Universal Robots PolyScope program: P1140 INVITE_Demo_1111.urp

Program P1140 INVITE_Demo_1111 (installation=default_INVITE directory=/programs createdIn=5.10.1 lastSavedIn=5.23.0 robotSerialNumber=20245590068)
Calibrated DH parameters: a=[0.00013, -0.03651, -0.389144, 0.000102, 0.000008, 0]; d=[0.162613, 192.230671, -179.915756, -12.181517, 0.099698, 0.099535]; alpha=[1.57038, 0.002205, 0.004138, 1.570804, -1.571025, 0]; deltaTheta=[-0.000001, 1.484886, 4.928506, -0.130209, 0, 0]
InitVariablesNode variables(variable(name=AMR_Position, expression=struct(position_identifier=0, x1=0, x2=0, y1=0, y2=0, theta1=0, theta2=0)), variable(name=CAM_Pose, expression=p[0,0,0,0,0,0]), variable(name=CAM_Relation, expression=""), variable(name=CMD_Abort, expression=False), variable(name=CMD_Clear, expression=False), variable(name=CMD_Reset, expression=False), variable(name=CMD_Start, expression=False), variable(name=CMD_Suspend, expression=False), variable(name=CMD_Unhold, expression=False), variable(name=CMD_Unsuspend, expression=False), variable(name=CNT_Rack_Output, expression=0), variable(name=FNC_Freedrive, expression=False), variable(name=PRC_TubCounter, expression=0), variable(name=PRC_TubNumber, expression=0), variable(name=STP, expression=0), variable(name=TMR_Barcode, expression=0), variable(name=easyPickCount, expression=0), variable(name=easyPickCount_5, expression=0), variable(name=easyPickNoObj, expression=0), variable(name=easyPickNoObj_5, expression=0), variable(name=easyPickParts, expression=0), variable(name=easyPickParts_5, expression=0))
BeforeStart
  Folder Scripts [hidden by the author, left out]
  Folder BeforeStarts [hidden by the author, left out]
  Script file /programs/04 Scripts/krish.script
    | def vibration_2():
    | 	set_analog_out(0,0.4)
    | 	sleep(0.8)
    | 	set_analog_out(0,0.0)
    | 	sleep(0.2)
    | end
    | 
    | def vibration_3():
    | 	set_analog_out(0,0.4)
    | 	sleep(0.7)
    | 	set_analog_out(0,0.0)
    | 	sleep(0.3)
    | end
    | 
    | def vibration_4():
    | 	set_analog_out(0,0.4)
    | 	sleep(0.6)
    | 	set_analog_out(0, 0.0)
    | 	sleep(0.5)
    | end
    | 
    | def vibration_1():
    | 	set_analog_out(0,0.4)
    | 	sleep(1)
    | 	set_analog_out(0,0.0)
    | 	sleep(0)
    | end
    | 
    | def move_tilt_in_steps(Pow_center, final_pose, steps):
    | 	i = 0
    | 	while i <= steps:
    | 		ratio = i / steps
    | 		pose_step = p[Pow_center[0] + ratio * (final_pose[0] - Pow_center[0]), Pow_center[1] + ratio * (final_pose[1] -Pow_center[1]),Pow_center[2] + ratio * (final_pose[2] - Pow_center[2]), Pow_center[3] + ratio * (final_pose[3] - Pow_center[3]), Pow_center[4] + ratio * (final_pose[4] - Pow_center[4]), Pow_center[5] + ratio * (final_pose[5] - Pow_center[5])]
    | 		movej(pose_step, a=1.2, v=0.15)
    | 		sleep(0.1)
    | 		i = i+1
    | 	end
    | end
    | 
    | def tilt_container(angle):
    | 	p_center = get_actual_tcp_pose()
    | 	hinge_offset = p[0,0,-0.23,0,0,0]
    | 	pivot_pose = pose_trans(p_center, hinge_offset)
    | 	pose_rel = pose_trans(pose_inv(pivot_pose), p_center)
    | 	angle_mid = (angle/2.0)*3.1416/180
    | 	angle_end = angle*3.1416/180
    | 	tilt_mid = p[0,0,0, -angle_mid, 0, 0]
    | 	tilt_end = p[0,0,0, -angle_end, 0, 0]
    | 	pose_rel_mid = pose_trans(tilt_mid, pose_rel)
    | 	pose_rel_end = pose_trans(tilt_end, pose_rel)
    | 	via_pose = pose_trans(pivot_pose, pose_rel_mid)
    | 	end_pose = pose_trans(pivot_pose, pose_rel_end)
    | 	movec(via_pose, end_pose, a=0.05, v=0.01, r=0.001)
    | 	p_center = get_actual_tcp_pose()
    | end
    | 
    | def deg2rad(d):
    | 	return d*3.141592/180
    | end
    | 
    | def map_tilt_to_ry_deg(container_deg):
    | 	#ry_deg = -0.875*container_deg +87.0
    | 	#return clamp(ry_deg, 5.0, 80.0)
    | 	if (Pow_name == "NaCl" or Pow_name == "Mannitol" or Pow_name == "CCS" or Pow_name == "lactose_loose"):
    | 		if ( level>=10.0):
    | 			ry_min = 10.0
    | 			ry_max = 75.0
    | 		elif (level<10.00 and level >1.00):
    | 			ry_min = 16.0
    | 			ry_max = 65.0
    | 		else:
    | 			ry_min=17.0
    | 			ry_max=75.0
    | 		end
    | 	else:
    | 		if ( level>=10.0):
    | 			ry_min = 0.0
    | 			ry_max = 55.0
    | 		elif (level<10.00 and level >1.00):
    | 			ry_min = 10.0
    | 			ry_max = 45.0
    | 		else:
    | 			ry_min=0.0
    | 			ry_max=50.0
    | 		end
    | 
    | 	end
    | 	local span_count = angle_max -angle_min
    | 	local span_ry = ry_max - ry_min
    | 
    | 	local t = (container_deg -angle_min)/span_count
    | 	local ry_deg = ry_max - t*span_ry
    | 
    | 	return clamp(ry_deg, ry_min, ry_max)
    | 
    | end
    | 
    | def caluclate_corrections(level):
    | 	z_high = 0.01
    | 	z_low = -0.08
    | 	y_high = -0.010
    | 	y_low = -0.03
    | 
    | 	scale = (level - 10.0) / (100.0-10.0)
    | 
    | 	global correction_z = z_low + scale*(z_high - z_low)
    | 	global correction_y = y_low + scale*(y_high -y_low)
    | 
    | end
    | 
    | def scoop_powder(p_center):
    | 	#lift_offset = p[0, 0, 0.05, 0, 0, 0]
    | 	vibration_voltage = 0.4
    | 	vibration_time = 3.0
    | 	diameter = 0.07
    | 	global scoop_radius_default = 0.0
    | 	#p_center = center_pose_t
    | 
    | 
    | 	if (level >=70.00):
    | 		approach_offset = p[0.008,0,0.22,0,0,0]
    | 		lift_offset = p[0, 0, 0.12, 0, 0, 0]
    | 		caluclate_corrections(level)
    | 	elif (level >=10.00 and level <70):
    | 		approach_offset = p[0.008,0,0.22,0,0,0]
    | 		lift_offset = p[0, 0, 0.15, 0, 0, 0]
    | 		caluclate_corrections(level)
    | 	elif (level<10.00 and level >= 1.00):
    | 		approach_offset = p[0.006,0,0.22,0,0,0]
    | 		correction_z = -0.08
    | 		correction_y = -0.01
    | 		lift_offset = p[0, 0, 0.14, 0, 0, 0]
    | 	else:
    | 		approach_offset = p[0.008,0,0.22,0,0,0]
    | 		correction_z = -0.08
    | 		correction_y = -0.01
    | 		lift_offset = p[0, 0, 0.14, 0, 0, 0]
    |  	end
    | 
    | 	if (spatula == "spatula_L"):
    | 		global spatula_depth = 0.015
    | 	elif (spatula == "spatula_M"):
    | 		global spatula_depth = 0.01
    | 	elif (spatula == "spatula_S"):
    | 		global spatula_depth = 0.006
    | 	elif (spatula == "spatula_flat_M"):
    | 		global spatula_depth = 0.001
    | 	elif (spatula == "spatula_flat_S"):
    | 		global spatula_depth = 0.005
    | 	end
    | 
    | 	scoop_radius_default = diameter/2 - spatula_depth
    | 	scoop_entry_pose = pose_trans(p_center, approach_offset)
    | 	movel(scoop_entry_pose, a=0.05, v=0.05)
    | 
    | 	scoop_start_rel = p[scoop_radius_default, 0, scoop_depth, 0, 0, 0]
    | 
    | 	rot_mid = p[0, 0, 0, 0, 0, 0.785]
    | 	rot_end = p[0, 0, 0, 0, 0, 1.5708]
    | 
    | 	scoop_via_rel = pose_trans(rot_mid, scoop_start_rel)
    | 	scoop_end_rel = pose_trans(rot_end, scoop_start_rel)
    | 
    | 	scoop_start_pose = pose_trans(p_center, scoop_start_rel)
    | 	scoop_via_pose = pose_trans(p_center, scoop_via_rel)
    | 	scoop_end_pose = pose_trans(p_center, scoop_end_rel)
    | 
    | 	movel(scoop_start_pose, a=0.3, v=0.7)
    | 
    | 	if (level<90.0):
    | 		Rotate()
    | 	end
    | 
    | 	#movec(scoop_via_pose, scoop_end_pose, a=0.03, v=0.05)
    | 	movec(scoop_via_pose, scoop_end_pose, a=0.03, v=0.02)
    | 	#movel(pose_trans(get_actual_tcp_pose(), p[0,0,0,0,0,deg2rad(90.0)]), a=0.03, v=0.05)
    | 	sleep(1.0)
    | 	local ry_deg = map_tilt_to_ry_deg(angle_deg)
    | 	local ry = deg2rad(ry_deg)
    | 	local end_rel = pose_trans(pose_inv(p_center), scoop_end_pose)
    | 	local end_rel_tilted = pose_trans(end_rel, p[0, 0, 0, 0, ry, 0])
    | 	global tilted_pose_in_base = pose_trans(p_center, p[0,correction_y,correction_z,end_rel_tilted[3],end_rel_tilted[4], end_rel_tilted[5]])
    | 	global tilted_pose_in_base = pose_trans(tilted_pose_in_base, p[0, 0, spatula_len, 0, 0, 0])
    | 
    | 	movel(tilted_pose_in_base, a=0.03, v=0.1)
    | 	set_analog_out(0, vibration_voltage)
    | 
    | 	local ry_level = deg2rad(ry_deg/1.5)
    | 	local end_rel_tilted_level = pose_trans(end_rel, p[0, 0, 0, 0, ry_level, 0])
    | 	local level_tilted_pose_in_base = pose_trans(p_center, p[0,correction_y,correction_z,end_rel_tilted_level[3],end_rel_tilted_level[4], end_rel_tilted_level[5]])
    | 	local level_tilted_pose_in_base = pose_trans(level_tilted_pose_in_base, p[0, 0, spatula_len, 0, 0, 0])
    | 
    | 	movel(level_tilted_pose_in_base, a=0.03, v=0.1)
    | 	#if (level>70.0):
    | 		#sleep(1.0)
    | 	#end
    | 	sleep(2.0)
    | 	#sleep(vibration_time)
    | 
    | 	movel(tilted_pose_in_base, a=0.03, v=0.1)
    | 	set_analog_out(0, 0.0)
    | 
    | 	tilt_pose_rel = pose_trans(pose_inv(p_center), tilted_pose_in_base)
    | 
    | 	lifted_pose_rel = pose_trans(lift_offset, tilt_pose_rel)
    | 
    | 	global lifted_pose = pose_trans(p_center, lifted_pose_rel)
    | 	movel(lifted_pose, a=0.03, v=0.1)
    | end
    | 
    | 
    | def center_pose():
    | 	trans_rel = p[-0.014, 0.06, -0.015, 0, 0, 0]
    | 
    | 	p_translated = pose_trans(place_pose, trans_rel)
    | 	cx = p_translated[0]
    | 	cy = p_translated[1]
    | 	cz = p_translated[2]
    | 
    | 	global p_center_vertical = p[cx,cy,cz, 0, 0, 4.08]
    | 
    | 	#movej(p_center_vertical, a =0.3, v =0.3)
    | 	return p_center_vertical
    | end
    | 
    | def updated_center_pose(p_center_vertical, angle_deg):
    | 	hinge_pose = pose_trans(p_center_vertical, p[0,0,-0.2,0,0,0])
    | 	local_rel = pose_trans(pose_inv(hinge_pose), p_center_vertical)
    | 
    | 	rot_tilt = p[0,0,0, -deg2rad(angle_deg),0,0]
    | 	local_rel_tilted = pose_trans(rot_tilt, local_rel)
    | 
    | 	global p_center = pose_trans(hinge_pose, local_rel_tilted)
    | 	return p_center
    | end
    | 
    | def tilt_send(angle):
    | 	socket_open("192.168.12.105", 80)
    | 	angle = 85.0 - angle
    | 	socket_send_string("Tilt,"+to_str(angle)+",0")
    | 	sync()
    | 	sleep(0.5)
    | 	socket_close()
    | end
    | 
    | def Motors_off():
    | 	socket_open("192.168.12.105", 80)
    | 	socket_send_string("Off,0,0")
    | 	sync()
    | 	sleep(0.5)
    | 	socket_close()
    | end
    | 
    | def Rotate():
    | 	socket_open("192.168.12.105", 80)
    | 	socket_send_string("FullRotation, 1, 2000")
    | 	sync()
    | 	sleep(0.5)
    | 	socket_close()
    | end
    | 
    | def tilt_to_home():
    | 	socket_open("192.168.12.105", 80)
    | 	socket_send_string("Home,0,0")
    | 	sync()
    | 	sleep(0.5)
    | 	socket_close()
    | end
  Script file /programs/04 Scripts/scooping.script
    | def scooping_init():
    | 	global W_EMPTY = 51.381
    | 	#global W_FULL = 300.010
    | 	global H_INNER = 0.15
    | 	global TCP_to_tip = 0.020
    | 	global depth_saftey = 0.005
    | 	global container_height = 0.120
    | 	global reach_margin = 0.03
    | 
    | 	global angle_min = 18.0
    | 	global angle_max = 68.0
    | 	global gain_per_percent = 0.5
    | 
    | 	global level_bias_below_center = 0.020
    | 
    | 	global level = 0.0
    | 	global tilt_angle_sent = 0.0
    | 	global w_dosed_total = 0.0
    | 	global last_scale = 0.0
    | 	global g_z0_hi = 0.01
    | 	global g_z100_hi = 0.14
    | 	global g_z_min = 0.030
    | 	global g_z_max = 0.150
    | 
    | 	#global g_exp = 0.80
    | 	#global g_k = 0.03
    | 	#global g_alpha = 0.7
    | 	global g_corr_max = 0.010
    | 
    | 	global g_prev_cum_w = -1.0
    | 	global g_depth_corr = 0.0
    | 	global spatula_len = 0.17
    | 	global target_g = 0.0
    | 	global scoop_ct = 0
    | 	global error_sum = 0.0
    | 	global error_sq_sum = 0.0
    | 	global scoop_g = 0.0
    | 
    | 	if (Pow_name=="NaCl"):
    | 		global W_FULL = 625.00
    | 		global g_exp = 0.80
    | 		global g_k = 0.03
    | 		global g_alpha = 0.7
    | 	elif (Pow_name == "Mannitol"):
    | 		global W_FULL = 300.00
    | 		global g_exp = 0.82
    | 		global g_k = 0.025
    | 		global g_alpha = 0.6
    | 	elif (Pow_name == "lactose_loose"):
    | 		global W_FULL = 250.0
    | 		global g_exp = 0.82
    | 		global g_k = 0.035
    | 		global g_alpha = 0.7
    | 	elif (Pow_name == "CCS"):
    | 		global W_FULL = 270.0
    | 		global g_exp = 0.82
    | 		global g_k = 0.035
    | 		global g_alpha = 0.7
    | 	elif (Pow_name == "Magnesium_sterate"):
    | 		global W_FULL = 220.0
    | 		global g_exp = 0.84
    | 		global g_k = 0.04
    | 		global g_alpha = 0.7
    | 	elif (Pow_name == "lactose_fine"):
    | 		global W_FULL = 330.0
    | 		global g_exp = 0.84
    | 		global g_k = 0.04
    | 		global g_alpha = 0.7
    | 	else:
    | 		popup("Unkwon powder type. Using default NaCl settings.", title="Calibration Warning")
    | 		global W_FULL = 300.0
    | 		global g_k = 0.03
    | 		global g_alpha = 0.7
    | 	end
    | 
    | 
    | end
    | 
    | def clamp(x, lo, hi):
    | 	if(x<lo):
    | 		return lo
    | 	elif (x>hi):
    | 		return hi
    | 	else:
    | 		return x
    | 	end
    | end
    | 
    | def compute_level_percent(W_now, weight_value):
    | 	local delta = weight_value - last_scale
    | 	if (delta<0.0):
    | 		delta = 0.0
    | 	end
    | 	global w_dosed_total = w_dosed_total + delta
    | 	global last_scale = weight_value
    | 
    | 	local W_eff = W_now-w_dosed_total
    | 	if (W_eff<W_EMPTY):
    | 		W_eff = W_EMPTY
    | 	end
    | 
    | 	level = 100.0* (W_eff -W_EMPTY)/ (W_FULL-W_EMPTY)
    | 	level = clamp(level,0.0,100.0)
    | 
    | 	#if (Task =="Emptying"):
    | 		#if (level>10.0):
    | 			#global spatula = "spatula_L"
    | 		#elif (level<=10.0 and level >1.0):
    | 			#global spatula = "spatula_M"
    | 		#else:
    | 			#global spatula = "spatula_S"
    | 		#end
    | 	#elif (Task == "Dosing"):
    | 		#if (level>10.0 and diff>=3.5):
    | 			#global spatula = "spatula_L"
    | 		#elif (level>10.0 and diff<3.5):
    | 			#global spatula = "spatula_M"
    | 		#elif (level<=10.0 and level >1.0):
    | 			#global spatula = "spatula_M"
    | 		#else:
    | 			#global spatula = "spatula_S"
    | 		#end
    | 	#end
    | 
    | 	return level
    | end
    | 
    | def compute_tilt_deg(level_percent):
    | 	angle = angle_min + gain_per_percent*(100.0-level_percent)
    | 	return clamp(angle, angle_min, angle_max)
    | 	#return angle
    | end
    | 
    | 
    | def tilt(level_percentage):
    | 	new_angle = compute_tilt_deg(level_percentage)
    | 	global angle_rel = new_angle - tilt_angle_sent
    | 
    | 	if my_abs(angle_rel)>2.0:
    | 		tilt_send(new_angle)
    | 		global angle_deg = new_angle
    | 		global tilt_angle_sent = new_angle
    | 		global p_center = updated_center_pose(p_center_vertical, angle_deg)
    | 	end
    | 
    | 	#if (level<85.0):
    | 		#tilt_send(angle_deg)
    | 	#end
    | end
    | 
    | def compute_scoop_depth(level, cum_w, target_g):
    | 	if (level >=10.0):
    | 		ratio = level/100.0
    | 		corrected = pow(ratio, g_exp)
    | 		base_z = g_z0_hi + (g_z100_hi - g_z0_hi)*corrected
    | 
    | 	elif (level<10.00 and level>=1.00):
    | 		z0 = 0.035
    | 		z100 = 0.140
    | 		ratio2 = level/100.0
    | 		base_z = z0 +(z100-z0)*ratio2
    | 	else:
    | 		base_z = 0.028
    | 	end
    | 
    | 	if (g_prev_cum_w<0):
    | 		g_prev_cum_w = cum_w
    | 
    | 	else:
    | 		global scoop_g = cum_w-g_prev_cum_w
    | 		g_prev_cum_w = cum_w
    | 
    | 		e = target_g -scoop_g
    | 
    | 		corr_proposed = g_k*e
    | 		g_depth_corr = (1.0 -g_alpha)*g_depth_corr + g_alpha*corr_proposed
    | 		g_depth_corr = clamp(g_depth_corr, -g_corr_max, g_corr_max)
    | 	end
    | 
    | 	z_tip = base_z - g_depth_corr
    | 	z_tip = clamp(z_tip, g_z_min, g_z_max)
    | 
    | 
    | 	return z_tip
    | end
    | 
    | def my_abs(val):
    | 	if (val<0):
    | 		return -val
    | 	else:
    | 		return val
    | 	end
    | end
    | 
    | 
    | def select_spatula(Pow_name, level, diff):
    | 	if (Pow_name == "lactose_fine" or Pow_name== "Magnesium_sterate"):
    | 		if (level >10.0):
    | 			return "spatula_flat_M"
    | 		else:
    | 			return "spatula_flat_s"
    | 		end
    | 
    | 	elif (Pow_name == "NaCl" and level >10.0 and diff>6.5):
    | 		return "spatula_L"
    | 	elif(Pow_name == "NaCl" and level> 10.0 and diff<=6.5):
    | 		return "spatula_M"
    | 	elif (Pow_name == "lactose_loose" and level >10.0 and diff>2.0):
    | 		return "spatula_L"
    | 	elif(Pow_name == "lactose_loose" and level> 10.0 and diff<=2.0):
    | 		return "spatula_M"
    | 	elif (Pow_name == "Mannitol" or Pow_name == "CCS" and level >10.0 and diff>3.2):
    | 		return "spatula_L"
    | 	elif(Pow_name == "Mannitol" or Pow_name == "CCS" and level> 10.0 and diff<=3.2):
    | 		return "spatula_M"
    | 	elif( level>1.0 and level <= 10.0):
    | 		return "spatula_M"
    | 	else:
    | 		return "spatula_S"
    | 	end
    | end
    | 
    | global target_g_table = [
    | 	"NaCl", "spatula_L", "6.5",
    | 	"NaCl", "spatula_M", "1.5",
    | 	"NaCl", "spatula_S", "0.135",
    | 
    | 	"Mannitol", "spatula_L", "2.85",
    | 	"Mannitol", "spatula_M", "0.8",
    | 	"Mannitol", "spatula_S", "0.075",
    | 
    | 	"CCS", "spatula_L", "2.45",
    | 	"CCS", "spatula_M", "0.6",
    | 	"CCS", "spatula_S", "0.075",
    | 
    | 	"lactose_loose", "spatula_L", "1.6",
    | 	"lactose_loose", "spatula_M", "0.5",
    | 	"lactose_loose", "spatula_S", "0.05",
    | 
    | 	"Magnesium_sterate", "spatula_flat_M", "0.5",
    | 	"Magnesium_sterate", "spatula_flat_S", "0.25",
    | 
    | 	"lactose_fine", "spatula_flat_M", "1.0",
    | 	"lactose_fine", "spatula_flat_S", "0.5"]
    | 
    | def get_target_g(Pow_name, spat_name):
    | 	local i = 0
    | 	local n = length(target_g_table)
    | 	while (i < n):
    | 		if (target_g_table[i] == Pow_name and target_g_table[i+1] == spat_name):
    | 			return to_num(target_g_table[i+2])
    | 		end
    | 		i = i+3
    | 	end
    | 	popup("No target_g match for: ", Pow_name, ", ", spatula)
    | 
    | end
    | def auto_tilt_and_scoop(W_now, target_weight, weight_value):
    | 	level = compute_level_percent(W_now, weight_value)
    | 
    | 	#global angle_deg = compute_tilt_deg(level)
    | 
    | 	#if(level>=10.0):
    | 		#target_g = 2.850
    | 	#elif(level<10.0 and level >=1.0):
    | 		#target_g= 0.8
    | 	#else:
    | 		#target_g = 0.060
    | 	#end
    | 
    | 
    | 	#if (Task =="Emptying"):
    | 		#if (level>10.0):
    | 			#target_g = 2.850
    | 		#elif (level<=10.0 and level >1.0):
    | 			#target_g = 0.8
    | 		#else:
    | 			#target_g = 0.060
    | 		#end
    | 	#elif (Task == "Dosing"):
    | 		#if (level>10.0 and diff>=3.5):
    | 			#target_g = 2.85
    | 		#elif (level>10.0 and diff<3.5):
    | 			#target_g = 0.8
    | 		#elif (level<=10.0 and level >1.0):
    | 			#target_g = 0.8
    | 		#else:
    | 			#target_g = 0.06
    | 		#end
    | 	#end
    | 
    | 	global spatula = select_spatula(Pow_name, level, diff)
    | 	global target_g = get_target_g(Pow_name, spatula)
    | 
    | 	global scoop_depth = compute_scoop_depth(level, weight_value, target_g)
    | 
    | 	tilt(level)
    | 	#p_center = get_actual_tcp_pose()
    | 
    | 	if (scoop_ct < 5 and g_prev_cum_w>0.0):
    | 		#local scoop_g = scoop_g
    | 		local error = target_g - scoop_g
    | 		error_sum = error_sum + error
    | 		error_sq_sum = error_sq_sum + error*error
    | 		scoop_ct = scoop_ct+1
    | 
    | 		if (scoop_ct==5):
    | 			local avg_error = error_sum/5.0
    | 			#local std_dev = sqrt(error_sq_sum/5.0) - (avg_error*avg_error))
    | 
    | 			if (my_abs(avg_error)>1.0):
    | 				g_k = 0.055
    | 				g_alpha = 0.85
    | 			elif (my_abs(avg_error)>0.6):
    | 				g_k= 0.045
    | 				g_alpha =0.75
    | 			elif (my_abs(avg_error)> 0.3):
    | 				g_k = 0.035
    | 				g_alpha = 0.65
    | 			elif (my_abs(avg_error)>0.1):
    | 				g_k = 0.025
    | 				g_alpha = 0.55
    | 			else:
    | 				g_k = 0.015
    | 				g_alpha = 0.45
    | 			end
    | 		end
    | 	end
    | 
    | 	scoop_powder(p_center)
    | end
    | 
    | 
    | def after_scoop():
    | 	tilt_send(angle_deg)
    | 	sleep(0.5)
    | 	movel(lifted_pose, a=0.05, v=0.2)
    | 	movel(tilted_pose_in_base, a=0.05, v=0.2)
    | 	set_analog_out(0,0.4)
    | 	movel(pose_trans(tilted_pose_in_base, p[-0.01,0,0,0,0,2.0]), a=0.05, v=0.2)
    | 	set_analog_out(0,0.0)
    | 	movel(lifted_pose, a=0.05, v=0.2)
    | 	tilt_to_home()
    | end
  Script file /programs/04 Scripts/dosing_pid.script
    | def dosing_pid(target_weight):
    | 	#kp = 0.005
    | 	#ki = 0.02
    | 	#kd = 0.2
    | 	#dt = 0.05
    | 	#current_error = 0.0
    | 	#Integral_error = 0.0
    | 	#previous_error = 0.0
    | 	#tilt_angle = -1.0
    | 	max_tilt_angle = -0.55
    | 	#current_pose = get_actual_tcp_pose()
    | 
    | 	while ( weight_value < target_weight and tilt_angle < max_tilt_angle):
    | 		weight_value = get_weight()
    | 		current_error = target_weight - weight_value
    | 		Integral_error = Integral_error + current_error*dt
    | 		derivative = (current_error - previous_error) / dt
    | 		tilt_increment = (kp * current_error) + (ki * Integral_error) + (kd * derivative)
    | 		current_pose = get_actual_tcp_pose()
    | 		tilt_angle = current_pose[4]
    | 		new_pose = pose_trans(current_pose, p[(tilt_increment/5), 0, 0, 0, tilt_increment, 0])
    | 		movel(new_pose, a = 0.075, v = 0.025, t = 0, r = 0)
    | 		previous_error = current_error
    | 		sleep(dt)
    | 	end
    | end
Robot Program (runOnlyOnce=false)
  Folder MAIN [hidden by the author, left out]
SubProgram -> Sub_Vision_V18
SubProgram  [hidden by the author, left out]
SubProgram -> Sub_Action_V4
